(* IEC 61131-3 sources: FibonacciChallenge/Class/SafetyCDIAS_Base (part 6) *)

          //Check for valid version
          if pPara^.aPara[1] = 0x01 then  //Version

            ret_code := READY;
            pResult^.aData[0] := 0x01;  //return version
            pResult^.aData[1]$UDINT := GetDiagVisualOffsetErrorCode();

            pResult^.uiLng := 12;

          else

            //invalid version, return error
            ret_code := 1$IprStates; //means iprStates::ERROR but a server error also exists

            pResult^.aData[0] := 0x0;
            pResult^.uiLng    := 4;

          end_if;

      end_case;
    else
      TRACE("(SafetyCDIAS_Base::GetDiagConnect::NewInst) Unknown command!");
      ret_code := 1$IprStates; //means iprStates::ERROR but a server error also exists

	END_CASE;

END_FUNCTION

FUNCTION VIRTUAL GLOBAL SafetyCDIAS_Base::FetchChannelInfo

  DiagVars.UserErrorInfoReady := FALSE;
  DiagVars.UserWantsErrorInfo := TRUE;

END_FUNCTION

FUNCTION VIRTUAL SafetyCDIAS_Base::GetChannelInfo
	VAR_INPUT
		pErrorMemUser 	: ^UINT;
		pErrorMem 	: ^USINT;
		ErrorDataLength 	: INT;
	END_VAR
	VAR_OUTPUT
		StateReady 	: BOOL;
	END_VAR
  VAR
  	i   : INT;
  END_VAR

  StateReady := DiagVars.UserErrorInfoReady;

  if StateReady then
    //copy error values in UserArray
    for i := 0 to ErrorDataLength-1 do

      pErrorMemUser^ := pErrorMem^;

      //set pointer to next entry
      pErrorMemUser += sizeof(UINT);
      pErrorMem += sizeof(USINT);
    end_for;
  end_if;

END_FUNCTION

FUNCTION VIRTUAL SafetyCDIAS_Base::GetDiagVisualOffsetErrorCode
	VAR_OUTPUT
		udOffset 	: UDINT;
	END_VAR

  //In the safety firmware for the CSCP and SCP there is only one byte for the errorcode
  //To have different errorcodes (between CSCP and SCP) the safetydesigner adds a fix offset of 1000 to the errorcodes of the SCP01x and SCP11x
  udOffset := 0;

END_FUNCTION
